Fanuc KAREL source: ka00053.KL

-- PROVISIONAL review KL for V1013-1; original PC SHA256 4a1214b371ff99f8e33b77a73381ea89f55638ee22255b11a702debbed738eb9
-- Incomplete behavior may be omitted. Consult companion uncertainty JSON. Do not deploy.
PROGRAM KA00053
%NOLOCKGROUP
-- UNRESOLVED_DECL SRC type=000101
-- UNRESOLVED_DECL DST type=000101
BEGIN
  -- UNRESOLVED_PC offsets 5-20; opcodes 49,4A
  -- UNRESOLVED_PC offsets 25-29; opcodes 7F
END KA00053
